Fanuc KAREL source: kt00368.KL

-- PROVISIONAL review KL for V940-1; original PC SHA256 028e514804d9adb8e251350913a18a8ea38d8fe2735be35947b14595e0ff28eb
-- Incomplete behavior may be omitted. Consult companion uncertainty JSON. Do not deploy.
PROGRAM KT00368
%NOLOCKGROUP
VAR
  I1 : INTEGER
  OUT : BOOLEAN
-- UNRESOLVED_DECL H2 type=002017
BEGIN
  -- V9_ZERO_TABLE_METADATA_HINT layout=0001; no indexed target words; source/name/runtime held
  -- UNRESOLVED_PC offsets 5-16; opcodes 2E,23
  -- UNRESOLVED_PC offsets 21-35; opcodes 2E,22,9D,33,B4
  -- UNRESOLVED_PC offsets 40-62; opcodes 21,22,9D,33,B3,5A,23
  -- UNRESOLVED_PC offsets 67-71; opcodes 7F
END KT00368
